(* IEC 61131-3 sources: codesys-washlet/codesys/src, 11 files *)

(* ---- E_WashAlarm.st ---- *)
(*
 * E_WashAlarm
 * 目的 : FB_Washlet が FAULT / ESTOP に入った理由（最初の1件だけ保持する）
 * 履歴 : 2026-10-30 新規作成
 *)
{attribute 'qualified_only'}  // CODESYS 拡張
{attribute 'strict'}          // CODESYS 拡張
TYPE E_WashAlarm :
(
    NONE                := 0,
    ESTOP_PRESSED       := 1,   (* 非常停止ボタンが押された（または配線が切れた） *)
    EXTEND_TIMEOUT      := 11,  (* ノズルが時間内に伸びきらない *)
    RETRACT_TIMEOUT     := 12,  (* ノズルが時間内に戻らない *)
    NOZZLE_SENSOR_BOTH  := 13,  (* 伸長端と収納端が同時に ON（センサ異常） *)
    WATER_OVER_TEMP     := 21,  (* 水温が上限を超えた。やけど防止 *)
    IO_LINK_LOST        := 31,  (* 機械（Web側）からの入力が途絶えた *)
    INVALID_STATE       := 99   (* CASE の ELSE。来てはいけない *)
);
END_TYPE

(* ---- E_WashState.st ---- *)
(*
 * E_WashState
 * 目的 : 温水洗浄便座コントローラ（FB_Washlet）の状態
 * 履歴 : 2026-10-30 新規作成
 *)
{attribute 'qualified_only'}  // CODESYS 拡張: E_WashState.IDLE の形でしか書けなくする
{attribute 'strict'}          // CODESYS 拡張: 列挙型に整数を直接代入できなくする
TYPE E_WashState :
(
    IDLE           := 0,   (* 待機。通常はノズル収納済み *)
    NOZZLE_EXTEND  := 1,   (* ノズル伸長中 *)
    SPRAY          := 2,   (* 噴射中 *)
    NOZZLE_RETRACT := 3,   (* ノズル収納中 *)
    ESTOP          := 10,  (* 非常停止中。動く出力はすべて OFF *)
    FAULT          := 20   (* 異常。リセット待ち *)
);
END_TYPE

(* ---- ST_WashInputs.st ---- *)
(*
 * ST_WashInputs
 * 目的 : 制御（FB_Washlet）が使う入力。変換層（FB_WashInputConv）が作る。
 *        中身は、構造体にする前の FB_Washlet の入力 9 本と同じ。
 *        生の値（ST_WashRawInputs）と違い、単位は換算済み、通信の健全性も判断済み。
 * 履歴 : 2026-11-06 新規作成（入力を構造体にまとめ、層に分けた）
 *)
TYPE ST_WashInputs :
STRUCT
    bEStopOk       : BOOL;   (* 非常停止が健全（NC接点。押される・断線で FALSE） *)
    bSeated        : BOOL;   (* 着座センサ *)
    bWashButton    : BOOL;   (* 「おしり」ボタン *)
    bStopButton    : BOOL;   (* 「止」ボタン（通常停止） *)
    bResetButton   : BOOL;   (* リセットボタン *)
    bNozzleAtFront : BOOL;   (* ノズル伸長端センサ *)
    bNozzleAtHome  : BOOL;   (* ノズル収納端センサ *)
    rWaterTemp     : REAL;   (* 水温 [℃] *)
    bIoHealthy     : BOOL;   (* 入力が生きている（通信ウォッチドッグ OK） *)
END_STRUCT
END_TYPE

(* ---- ST_WashOutputs.st ---- *)
(*
 * ST_WashOutputs
 * 目的 : 機械を動かす出力（アクチュエータ）4 つ。
 *        状態を知らせる出力（eState・eAlarm・許可）はここに入れない。
 *        「機械を動かす出力」と「状態を知らせる出力」を分けるため。
 * 履歴 : 2026-11-06 新規作成（出力を構造体にまとめ、層に分けた）
 *)
TYPE ST_WashOutputs :
STRUCT
    bNozzleExtend  : BOOL;   (* ノズル伸長 *)
    bNozzleRetract : BOOL;   (* ノズル収納 *)
    bPump          : BOOL;   (* 噴射ポンプ *)
    bHeater        : BOOL;   (* 温水ヒーター *)
END_STRUCT
END_TYPE

(* ---- ST_WashRawInputs.st ---- *)
(*
 * ST_WashRawInputs
 * 目的 : IO から来る「生の値」。I/O 層（PRG_IoModbus）が詰め、変換層（FB_WashInputConv）が読む。
 *        実機の IO ユニットに替えるときは、この構造体に I/O マッピングで値を入れる。
 *        単位の換算や判断はしない。来た値をそのまま持つ。
 * 履歴 : 2026-11-06 新規作成（入力を構造体にまとめ、層に分けた）
 *)
TYPE ST_WashRawInputs :
STRUCT
    bEStopOk       : BOOL;   (* 非常停止 NC接点。閉 = TRUE = 健全 *)
    bSeated        : BOOL;   (* 着座センサ *)
    bWashButton    : BOOL;   (* 「おしり」ボタン *)
    bStopButton    : BOOL;   (* 「止」ボタン *)
    bResetButton   : BOOL;   (* リセットボタン *)
    bNozzleAtFront : BOOL;   (* ノズル伸長端センサ *)
    bNozzleAtHome  : BOOL;   (* ノズル収納端センサ *)
    wWaterTempRaw  : WORD;   (* 水温 [℃×100]（38.00℃ → 3800） *)
    wHeartbeat     : WORD;   (* 機械側のハートビート。毎回 +1 される *)
END_STRUCT
END_TYPE

(* ---- GVL_IO.st ---- *)
(*
 * GVL_IO
 * 目的 : 層と層の受け渡しの置き場所。ロジックは %IX/%QX や Modbus 配列を直接使わず、ここを使う。
 *
 *   stRawIn  … I/O 層（PRG_IoModbus.ReadInputs）が書く。IO から来た生の値
 *   stIn     … 変換層（FB_WashInputConv）の出力を PLC_PRG が書く。制御が使う値
 *   stOut    … 制御層（FB_Washlet）の出力を PLC_PRG が書く
 *   stRawOut … PLC_PRG が stOut をコピーして書く。I/O 層（PRG_IoModbus.WriteOutputs）が読む
 *
 * 各変数を書くのは 1 か所だけ。
 * 実機の IO ユニットに替えるときは、stRawIn / stRawOut を I/O マッピング先にして、
 * PRG_IoModbus を外すだけで済む（変換層と制御層はそのまま）。
 *
 * 履歴 : 2026-10-30 新規作成
 *        2026-11-06 個別の BOOL をやめ、構造体 4 つにした
 *)
VAR_GLOBAL
    stRawIn  : ST_WashRawInputs;   (* 入力：IO → PLC（生の値） *)
    stIn     : ST_WashInputs;      (* 入力：制御が使う値 *)
    stOut    : ST_WashOutputs;     (* 出力：制御の結果 *)
    stRawOut : ST_WashOutputs;     (* 出力：PLC → IO *)
END_VAR

(* ---- GVL_Modbus.st ---- *)
(*
 * GVL_Modbus
 * 目的 : Web 側の「機械（plant）」とのやり取り（Modbus TCP）
 *   aFromTS : Holding Register（TS → PLC）＝ 機械のセンサ・ボタン
 *   aToTS   : Input Register  （PLC → TS）＝ PLC の出力・状態
 * レジスタの中身は README のレジスタマップ表を参照。
 * Modbus TCP Slave Device の I/O マッピングで、この2つの配列に割り当てる。
 * 履歴 : 2026-10-30 新規作成
 *        2026-10-30 機械モデルを Web 側に移したので、10 ワードずつに整理
 *)
VAR_GLOBAL
    aFromTS : ARRAY[0..9] OF WORD;
    aToTS   : ARRAY[0..9] OF WORD;
END_VAR

(* ---- FB_WashInputConv.st ---- *)
(*
 * FB_WashInputConv
 * 目的 : 変換層。IO から来た生の値（ST_WashRawInputs）を、制御が使う値（ST_WashInputs）にする。
 *        - 水温の換算 [℃×100] → [℃]
 *        - 通信ウォッチドッグ（ハートビートが T_LINK_TIMEOUT の間変わらなければ、入力を信用しない）
 *        IO の種類（Modbus か、実機の IO ユニットか）には関係しない。差し替えても、ここはそのまま使う。
 *
 * 入力:
 *   stRawIn   IO から来た生の値
 * 出力:
 *   stIn      制御が使う値
 *
 * 履歴 : 2026-11-06 新規作成（PLC_PRG にあった換算とウォッチドッグを移した）
 *)
FUNCTION_BLOCK FB_WashInputConv
VAR_INPUT
    stRawIn : ST_WashRawInputs;
END_VAR
VAR_OUTPUT
    stIn : ST_WashInputs;
END_VAR
VAR
    tonLinkLost : TON;
    wLastBeat   : WORD;   (* 前のサイクルに見えたハートビート *)
END_VAR
VAR CONSTANT
    T_LINK_TIMEOUT : TIME := T#500MS;   (* Web 側の書き込み周期 50 ms の 10 倍 *)
    R_TEMP_SCALE   : REAL := 100.0;     (* [℃×100] → [℃] *)
END_VAR

(* ---- 1. ボタン・センサ ---- *)
// チャタリング除去を入れるなら、ここ（ボタンやセンサごとに TON / TOF をかける）。
// 今は Web 側の機械モデルなので、接点のばたつきが無く、入れていない。
stIn.bEStopOk       := stRawIn.bEStopOk;
stIn.bSeated        := stRawIn.bSeated;
stIn.bWashButton    := stRawIn.bWashButton;
stIn.bStopButton    := stRawIn.bStopButton;
stIn.bResetButton   := stRawIn.bResetButton;
stIn.bNozzleAtFront := stRawIn.bNozzleAtFront;
stIn.bNozzleAtHome  := stRawIn.bNozzleAtHome;

(* ---- 2. 水温の換算 ---- *)
stIn.rWaterTemp := WORD_TO_REAL(stRawIn.wWaterTempRaw) / R_TEMP_SCALE;   (* [℃] *)

(* ---- 3. 通信ウォッチドッグ ---- *)
// ハートビートが止まったら、センサの値は「最後に見えた値」でしかない。信用しない。
// TON は毎サイクル呼ぶ（IF の中に入れない）
tonLinkLost(IN := stRawIn.wHeartbeat = wLastBeat, PT := T_LINK_TIMEOUT);
wLastBeat := stRawIn.wHeartbeat;
stIn.bIoHealthy := NOT tonLinkLost.Q;

(* ---- FB_Washlet.st ---- *)
(*
 * FB_Washlet
 * 目的 : 温水洗浄便座のノズル・ポンプ・ヒーターを制御する。
 *        非常停止とインターロックの学習用サンプル。
 *
 * 考え方（優先順位の高い順）:
 *   1. 非常停止 … どの状態からでも ESTOP へ。動く出力はすべて OFF。
 *                  解除しただけでは動かない。リセット操作が必要。
 *   2. 異常      … センサ矛盾・水温上限・タイムアウトで FAULT へ。
 *   3. インターロック … 「条件がそろわないと、その動作をさせない」。
 *                  状態遷移と出力の両方でチェックする（二重化）。
 *
 * ※ 本物の非常停止は、ソフトではなく安全リレー／安全PLCで
 *    動力を物理的に切る。この FB は「通常PLC側の振る舞い」の学習用。
 *
 * 入力:
 *   stIn            制御が使う入力（ST_WashInputs。中身は構造体の宣言を参照）
 *                   VAR_INPUT（値渡し）にしている理由:
 *                   - 数十バイトと小さく、コピーの重さは気にならない
 *                   - FB を呼んだ時点の値がコピーされ、1 サイクルの間は値が変わらない
 *                   - モニタで、FB が判断に使った値そのものが見える
 * 出力（機械を動かす出力）:
 *   stOut           ノズル伸長・収納、噴射ポンプ、温水ヒーター（ST_WashOutputs）
 * 出力（状態を知らせる出力。機械は動かさない）:
 *   eState / eAlarm                 状態と、最初に起きた異常
 *   bExtendPermit / bSprayPermit    インターロック成立（監視用）
 *
 * 履歴 : 2026-10-30 新規作成
 *        2026-11-06 入力 9 本を stIn 1 本に、アクチュエータの出力を stOut にまとめた（ロジックは変えていない）
 *)
FUNCTION_BLOCK FB_Washlet
VAR_INPUT
    stIn : ST_WashInputs;
END_VAR
VAR_OUTPUT
    stOut          : ST_WashOutputs;
    eState         : E_WashState := E_WashState.IDLE;
    eAlarm         : E_WashAlarm := E_WashAlarm.NONE;
    bExtendPermit  : BOOL;
    bSprayPermit   : BOOL;
END_VAR
VAR
    rtrigWash   : R_TRIG;
    rtrigReset  : R_TRIG;
    tonExtend   : TON;
    tonRetract  : TON;
    tonSpray    : TON;
    bTempOk     : BOOL;
    bHeatDemand : BOOL;   (* ヒーターのヒステリシス保持 *)
END_VAR
VAR CONSTANT
    T_EXTEND_TIMEOUT  : TIME := T#3S;    (* 設計値。実機に合わせて調整 *)
    T_RETRACT_TIMEOUT : TIME := T#3S;
    T_SPRAY_MAX       : TIME := T#60S;   (* 押しっぱなし防止の自動停止 *)
    R_TEMP_MAX        : REAL := 42.0;    (* [℃] これ以上は噴射させない *)
    R_TEMP_TARGET     : REAL := 38.0;    (* [℃] ヒーター目標 *)
    R_TEMP_HYST       : REAL := 1.0;     (* [℃] ヒーターのON/OFF幅 *)
END_VAR

(* ---- 1. FB は毎サイクル呼ぶ（IN で制御する） ---- *)
rtrigWash(CLK := stIn.bWashButton);
rtrigReset(CLK := stIn.bResetButton);
tonExtend (IN := eState = E_WashState.NOZZLE_EXTEND,  PT := T_EXTEND_TIMEOUT);
tonRetract(IN := eState = E_WashState.NOZZLE_RETRACT, PT := T_RETRACT_TIMEOUT);
tonSpray  (IN := eState = E_WashState.SPRAY,          PT := T_SPRAY_MAX);

(* ---- 2. インターロック条件 ---- *)
bTempOk       := stIn.rWaterTemp < R_TEMP_MAX;
bExtendPermit := stIn.bEStopOk AND stIn.bIoHealthy AND stIn.bSeated AND stIn.bNozzleAtHome AND bTempOk;
bSprayPermit  := stIn.bEStopOk AND stIn.bIoHealthy AND stIn.bSeated AND stIn.bNozzleAtFront AND bTempOk;

(* ---- 3. 非常停止・異常の割り込み（CASE より先に判定する） ---- *)
IF NOT stIn.bEStopOk THEN
    IF eState <> E_WashState.ESTOP THEN
        eState := E_WashState.ESTOP;
        IF eAlarm = E_WashAlarm.NONE THEN
            eAlarm := E_WashAlarm.ESTOP_PRESSED;
        END_IF
    END_IF
ELSIF eState <> E_WashState.ESTOP AND eState <> E_WashState.FAULT THEN
    IF NOT stIn.bIoHealthy THEN
        // 入力が止まったら、センサの値は「最後に見えた値」でしかない。信用せず止める
        eState := E_WashState.FAULT;
        eAlarm := E_WashAlarm.IO_LINK_LOST;
    ELSIF stIn.bNozzleAtFront AND stIn.bNozzleAtHome THEN
        eState := E_WashState.FAULT;
        eAlarm := E_WashAlarm.NOZZLE_SENSOR_BOTH;
    ELSIF NOT bTempOk THEN
        eState := E_WashState.FAULT;
        eAlarm := E_WashAlarm.WATER_OVER_TEMP;
    END_IF
END_IF

(* ---- 4. 通常の状態遷移 ---- *)
CASE eState OF
E_WashState.IDLE:
    IF NOT stIn.bNozzleAtHome THEN
        eState := E_WashState.NOZZLE_RETRACT;      // 起動時など、出ていたら先に戻す
    ELSIF rtrigWash.Q AND bExtendPermit THEN
        eState := E_WashState.NOZZLE_EXTEND;
    END_IF

E_WashState.NOZZLE_EXTEND:
    IF NOT stIn.bSeated OR stIn.bStopButton THEN
        eState := E_WashState.NOZZLE_RETRACT;
    ELSIF stIn.bNozzleAtFront THEN
        eState := E_WashState.SPRAY;
    ELSIF tonExtend.Q THEN
        eState := E_WashState.FAULT;
        eAlarm := E_WashAlarm.EXTEND_TIMEOUT;
    END_IF

E_WashState.SPRAY:
    IF NOT bSprayPermit OR stIn.bStopButton OR tonSpray.Q THEN
        eState := E_WashState.NOZZLE_RETRACT;      // 離席・止・時間切れは「正常な停止」
    END_IF

E_WashState.NOZZLE_RETRACT:
    IF stIn.bNozzleAtHome THEN
        eState := E_WashState.IDLE;
    ELSIF tonRetract.Q THEN
        eState := E_WashState.FAULT;
        eAlarm := E_WashAlarm.RETRACT_TIMEOUT;
    END_IF

E_WashState.ESTOP:
    // 解除しただけでは動かさない。解除＋リセット操作で、安全側（収納）から再開
    IF stIn.bEStopOk AND rtrigReset.Q THEN
        eAlarm := E_WashAlarm.NONE;
        eState := E_WashState.NOZZLE_RETRACT;
    END_IF

E_WashState.FAULT:
    // 原因が残っているうちはリセットを受け付けない
    IF rtrigReset.Q AND stIn.bIoHealthy AND bTempOk AND NOT (stIn.bNozzleAtFront AND stIn.bNozzleAtHome) THEN
        eAlarm := E_WashAlarm.NONE;
        eState := E_WashState.NOZZLE_RETRACT;
    END_IF

ELSE
    eState := E_WashState.FAULT;
    eAlarm := E_WashAlarm.INVALID_STATE;
END_CASE

(* ---- 5. ヒーターのヒステリシス ---- *)
IF stIn.rWaterTemp < R_TEMP_TARGET - R_TEMP_HYST THEN
    bHeatDemand := TRUE;
ELSIF stIn.rWaterTemp >= R_TEMP_TARGET THEN
    bHeatDemand := FALSE;
END_IF

(* ---- 6. 出力（書き込みはここだけ）。状態に加えて条件をもう一度かける ---- *)
stOut.bNozzleExtend  := eState = E_WashState.NOZZLE_EXTEND  AND stIn.bEStopOk AND stIn.bSeated;
stOut.bNozzleRetract := eState = E_WashState.NOZZLE_RETRACT AND stIn.bEStopOk AND stIn.bIoHealthy;
stOut.bPump          := eState = E_WashState.SPRAY          AND bSprayPermit;
stOut.bHeater        := bHeatDemand AND stIn.bEStopOk AND stIn.bIoHealthy AND bTempOk
                  AND eState <> E_WashState.FAULT
                  AND eState <> E_WashState.ESTOP;   // 解除しただけでは何も動かさない（ヒーターも）

(* ---- PLC_PRG.st ---- *)
(*
 * PLC_PRG
 * 目的 : 層を順に呼ぶ。
 *        I/O 層（入力）→ 変換層 → 制御層 → 出力のコピー → I/O 層（出力）
 *
 *   I/O 層  : PRG_IoModbus      Modbus 配列 ⇔ GVL_IO.stRawIn / stRawOut
 *   変換層  : FB_WashInputConv  生の値 → 制御が使う値（換算・通信ウォッチドッグ）
 *   制御層  : FB_Washlet        判断（非常停止・異常・インターロック・状態遷移）
 *
 * GVL_IO の各変数を書くのは 1 か所だけ（stRawIn は PRG_IoModbus、ほかはここ）。
 *
 * 構成 : 機械（ノズル・ヒーター・温度センサ・ボタン・非常停止）は Web 側にある。
 *        PLC は Modbus で「センサを読んで、出力を返す」だけ。実機の PLC と同じ立場。
 *        実機の IO ユニットに替えるときは、I/O 層だけを替える。
 *
 * 履歴 : 2026-10-30 新規作成
 *        2026-10-30 PRG_Sim を廃止。機械モデルを Web 側に移した
 *        2026-11-06 層に分けた。詰め替えを PRG_IoModbus、換算とウォッチドッグを FB_WashInputConv へ移した
 *)
PROGRAM PLC_PRG
VAR
    fbInputConv : FB_WashInputConv;
    fbWashlet   : FB_Washlet;
END_VAR

(* ---- 1. I/O 層（入力）：aFromTS → GVL_IO.stRawIn ---- *)
PRG_IoModbus.ReadInputs();

(* ---- 2. 変換層：生の値 → 制御が使う値 ---- *)
fbInputConv(stRawIn := GVL_IO.stRawIn);
GVL_IO.stIn := fbInputConv.stIn;

(* ---- 3. 制御層 ---- *)
fbWashlet(stIn := GVL_IO.stIn);
GVL_IO.stOut := fbWashlet.stOut;

(* ---- 4. 出力のコピー ---- *)
// 実機で出力の向き（反転など）を合わせるなら、ここで詰め替える。今はそのまま
GVL_IO.stRawOut := GVL_IO.stOut;

(* ---- 5. I/O 層（出力）：GVL_IO.stRawOut と状態 → aToTS ---- *)
PRG_IoModbus.eState        := fbWashlet.eState;
PRG_IoModbus.eAlarm        := fbWashlet.eAlarm;
PRG_IoModbus.bExtendPermit := fbWashlet.bExtendPermit;
PRG_IoModbus.bSprayPermit  := fbWashlet.bSprayPermit;
PRG_IoModbus.WriteOutputs();

(* ---- PRG_IoModbus.st ---- *)
(*
 * PRG_IoModbus
 * 目的 : I/O 層。Modbus の配列と GVL_IO の生の値を、相互に詰め替える。
 *        今は Web 側の機械モデルと Modbus TCP でつないでいるので、この PRG がある。
 *        実機の IO ユニットに替えるときは、この PRG を外し、
 *        GVL_IO.stRawIn / stRawOut を I/O マッピングで割り当てる。
 *
 * 呼び方（PLC_PRG から）:
 *   PRG_IoModbus.ReadInputs();    サイクルの最初。aFromTS → GVL_IO.stRawIn
 *   PRG_IoModbus.WriteOutputs();  サイクルの最後。GVL_IO.stRawOut と状態 → aToTS
 *
 * 入力（WriteOutputs の前に PLC_PRG が入れる。画面に出す状態。機械は動かさない）:
 *   eState / eAlarm                 状態と、最初に起きた異常
 *   bExtendPermit / bSprayPermit    インターロック成立
 *
 * レジスタの並びは README のレジスタマップ表のとおり（構造体にする前から変えていない）。
 *
 * 履歴 : 2026-11-06 新規作成（PLC_PRG にあった Modbus の詰め替えを移した）
 *)
PROGRAM PRG_IoModbus
VAR_INPUT
    eState        : E_WashState;
    eAlarm        : E_WashAlarm;
    bExtendPermit : BOOL;
    bSprayPermit  : BOOL;
END_VAR
VAR
    wInBits    : WORD;   (* HR0 のビット。画面へのエコーにも使う *)
    wOutBits   : WORD;
    wEchoBits  : WORD;
    wHeartbeat : WORD;   (* PLC 側のハートビート *)
END_VAR

(* 本体は使わない。ReadInputs / WriteOutputs を呼ぶ *)

ACTION ReadInputs
(* ---- 機械 → PLC：aFromTS → GVL_IO.stRawIn ---- *)
wInBits := GVL_Modbus.aFromTS[0];
GVL_IO.stRawIn.bEStopOk       := wInBits.0;   (* 接点が閉じている = 1 = 健全 *)
GVL_IO.stRawIn.bSeated        := wInBits.1;
GVL_IO.stRawIn.bWashButton    := wInBits.2;
GVL_IO.stRawIn.bStopButton    := wInBits.3;
GVL_IO.stRawIn.bResetButton   := wInBits.4;
GVL_IO.stRawIn.bNozzleAtFront := wInBits.5;
GVL_IO.stRawIn.bNozzleAtHome  := wInBits.6;
GVL_IO.stRawIn.wWaterTempRaw  := GVL_Modbus.aFromTS[1];   (* [℃×100] のまま。換算は変換層 *)
GVL_IO.stRawIn.wHeartbeat     := GVL_Modbus.aFromTS[2];
END_ACTION

ACTION WriteOutputs
(* ---- PLC → 機械：GVL_IO.stRawOut → aToTS ---- *)
wOutBits := 0;
wOutBits.0 := GVL_IO.stRawOut.bNozzleExtend;
wOutBits.1 := GVL_IO.stRawOut.bNozzleRetract;
wOutBits.2 := GVL_IO.stRawOut.bPump;
wOutBits.3 := GVL_IO.stRawOut.bHeater;
wOutBits.4 := bExtendPermit;
wOutBits.5 := bSprayPermit;

(* PLC から見えている入力を、そのまま返す（画面の「PLC の気持ち」用） *)
wEchoBits := wInBits;
wEchoBits.7 := GVL_IO.stIn.bIoHealthy;

wHeartbeat := wHeartbeat + 1;

GVL_Modbus.aToTS[0] := TO_WORD(eState);
GVL_Modbus.aToTS[1] := TO_WORD(eAlarm);
GVL_Modbus.aToTS[2] := wOutBits;
GVL_Modbus.aToTS[3] := wEchoBits;
GVL_Modbus.aToTS[4] := GVL_IO.stRawIn.wWaterTempRaw;   (* PLC が受け取った水温 [℃×100] *)
GVL_Modbus.aToTS[5] := wHeartbeat;
END_ACTION

END_PROGRAM
